FUNCTION_BLOCK FINAL SEQ_ModuleSequence EXTENDS GEN_Sequence
VAR_IN_OUT
    DevList : ST_ControlModuleDevList;
END_VAR
VAR
END_VAR

SUPER^();

METHOD PRIVATE InitAlarms : BOOL
END_METHOD

METHOD PRIVATE RaiseAlarm : BOOL
VAR_INPUT
	AlarmId : UDINT;
END_VAR
CASE AlarmId OF
0:
	;
END_CASE
END_METHOD

METHOD PROTECTED RunSteps
Steps();
END_METHOD

ACTION Steps:
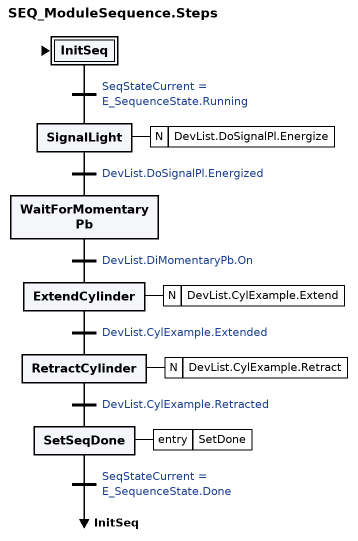
INITIAL_STEP InitSeq:
END_STEP
TRANSITION FROM InitSeq TO SignalLight
    := SeqStateCurrent = E_SequenceState.Running;
END_TRANSITION
STEP SignalLight:
    DevList.DoSignalPl.Energize(N);
END_STEP
TRANSITION FROM SignalLight TO WaitForMomentaryPb
    := DevList.DoSignalPl.Energized;
END_TRANSITION
STEP WaitForMomentaryPb:
END_STEP
TRANSITION FROM WaitForMomentaryPb TO ExtendCylinder
    := DevList.DiMomentaryPb.On;
END_TRANSITION
STEP ExtendCylinder:
    DevList.CylExample.Extend(N);
END_STEP
TRANSITION FROM ExtendCylinder TO RetractCylinder
    := DevList.CylExample.Extended;
END_TRANSITION
STEP RetractCylinder:
    DevList.CylExample.Retract(N);
END_STEP
TRANSITION FROM RetractCylinder TO SetSeqDone
    := DevList.CylExample.Retracted;
END_TRANSITION
STEP SetSeqDone:
    SetDone(P1);  // entry action
END_STEP
TRANSITION FROM SetSeqDone TO InitSeq
    := SeqStateCurrent = E_SequenceState.Done;
END_TRANSITION
END_ACTION

END_FUNCTION_BLOCK

(* stored: Version 1.1.0.1, ProductVersion 3.1.4024.12
   POU SEQ_ModuleSequence: Id {8d99d55f-7e79-41e9-a1b4-612faf9c000b}, SpecialFunc None
   Folder Override Methods: Id {1edc1085-d9e2-42dc-960b-f97ab143976d}
   Method InitAlarms: Id {c81da89c-fffe-4986-b286-fc43c7a28874}
   Method RaiseAlarm: Id {4d22e97d-7f12-40a0-9a3e-7314c8b752ce}
   Method RunSteps: Id {09379d0e-678f-4d9b-a369-46ffd832bc07}
   Action Steps: Id {34b69fa3-68f5-404c-90f2-a0917d99fb99} *)
